Staubli VAL3: stop.pgx

program stop()
// Safe stop routine: halts motion and resets feeder valve without dropping held parts.
begin
  resetMotion()
  bOut10 = false
  putln("Lab2B stopped safely - gripper state preserved")
end
